Fanuc KAREL source: kt00534.KL

-- PROVISIONAL review KL for V940-1; original PC SHA256 604769a4f6045d0a4059e6bb614d87e053f6346bad337882f98a676199e69df3
-- Incomplete behavior may be omitted. Consult companion uncertainty JSON. Do not deploy.
PROGRAM KT00534
%NOLOCKGROUP
-- UNRESOLVED_DECL P1 type=000199
-- UNRESOLVED_DECL P2 type=000101
-- UNRESOLVED_DECL OUT type=000101
BEGIN
  -- V9_ZERO_TABLE_METADATA_HINT layout=0001; no indexed target words; source/name/runtime held
  -- UNRESOLVED_PC offsets 5-34; opcodes 49,7E,49,60,4A
  -- UNRESOLVED_PC offsets 39-43; opcodes 7F
END KT00534
